TYPE "ST_TwoHandDevice"
VERSION : 0.1
   STRUCT
      Armed : Bool;
      SafeActive : Bool;
      SafePrevious : Bool;
      StartPulse : Bool;
   END_STRUCT;

END_TYPE

